(* IEC 61131-3 sources: plc-st-coding-agent/progress/evidence/f14_v14_remaining_20261113/jobs/codex_minimax-m27 (part 6) *)

(* ---- self-hard-07.candidate_01.st ---- *)
FUNCTION_BLOCK FB
VAR_INPUT
    mode                : INT;
    resetBtn            : BOOL;
    scanSeconds         : REAL;
    tempSP              : REAL;
    tempPV              : REAL;
    flowPV              : REAL;
    manualFlowSP        : REAL;
    manualValve         : REAL;
END_VAR
VAR_OUTPUT
    flowSP              : REAL;
    valveCommand        : REAL;
    fault               : BOOL;
    normalMode          : BOOL;
END_VAR
VAR
    accT                : REAL := 0.0;
    accF                : REAL := 0.0;
    mode_prev           : INT := 999;
    prev_resetBtn       : BOOL := FALSE;
    first_scan          : BOOL := TRUE;
END_VAR
VAR_TEMP
    eT                  : REAL;
    eF                  : REAL;
    trial               : REAL;
    reset_rising        : BOOL;
    mode_changed        : BOOL;
END_VAR
(* ENGINEERING_CONTRACT
 * =============================================================================
 * Modes: 0=Manual(FB), 1=Auto(inner PI), 2=Cascade(both PI loops)
 * Normal operation: mode in {0,1,2}, 0 < scanSeconds <= 10.0
 * Fault: mode outside {0,1,2} OR scanSeconds <= 0 OR scanSeconds > 10
 * -----------------------------------------------------------------------------
 * Output state retention (per LTL spec):
 * - Mode switch to 2 (cascade): flowSP, valveCommand HOLD prev; normalMode=FALSE
 * - Mode switch to 0/1: flowSP=manualFlowSP, valveCommand HOLD prev; normalMode=FALSE
 * - Manual (mode=0) normal cycle: flowSP=manualFlowSP, valveCommand=manualValve
 * - Auto (mode=1) normal cycle: flowSP=manualFlowSP; valveCommand=PI(clamped)
 * - Cascade (mode=2) normal cycle: flowSP=PI(clamped), valveCommand=PI(clamped)
 * - Fault: flowSP=manualFlowSP, valveCommand=manualValve, normalMode=FALSE
 * - Reset rising edge: same as fault initialization, fault still reports truthfully
 * -----------------------------------------------------------------------------
 * Integrators (anti-windup back-calculation):
 * - accT unit: t/h; accF unit: %; both pre-set to 0 on reset/fault/first scan
 * - acc update after output limit: acc = limited_output - Kp*e
 * - On mode change to cascade, both accT and accF retain prior cycle values
 * -----------------------------------------------------------------------------
 * Timing: Ki defined per second; scanSeconds multiplied explicitly
 * Boundaries: flowSP [0,50] t/h; valveCommand [0,100] %
 * =============================================================================
 *)
(* CONTRACT_RULES [] *)

reset_rising := resetBtn AND NOT prev_resetBtn;
mode_changed := (mode <> mode_prev);

fault := (mode < 0) OR (mode > 2) OR (scanSeconds <= 0.0) OR (scanSeconds > 10.0);

IF first_scan OR reset_rising THEN
    flowSP := manualFlowSP;
    valveCommand := manualValve;
    accT := 0.0;
    accF := 0.0;
    normalMode := FALSE;
    first_scan := FALSE;
ELSIF fault THEN
    flowSP := manualFlowSP;
    valveCommand := manualValve;
    accT := 0.0;
    accF := 0.0;
    normalMode := FALSE;
ELSE
    IF mode_changed THEN
        normalMode := FALSE;
        IF mode = 2 THEN
            // Cascade: hold both outputs
            // accT, accF retained for bumpless entry
        ELSIF (mode = 0) OR (mode = 1) THEN
            flowSP := manualFlowSP;
            // valveCommand held
        END_IF;
    ELSE
        normalMode := TRUE;
        IF mode = 2 THEN
            // Outer loop PI
            eT := tempSP - tempPV;
            accT := accT + 0.2 * eT * scanSeconds;
            trial := accT + 0.2 * eT * scanSeconds;
            flowSP := 1.0 * eT + trial;
            flowSP := LIMIT(0.0, flowSP, 50.0);
            accT := flowSP - 1.0 * eT;
            // Inner loop PI
            eF := flowSP - flowPV;
            accF := accF + 0.5 * eF * scanSeconds;
            trial := accF + 0.5 * eF * scanSeconds;
            valveCommand := 2.0 * eF + trial;
            valveCommand := LIMIT(0.0, valveCommand, 100.0);
            accF := valveCommand - 2.0 * eF;
        ELSIF mode = 1 THEN
            // Auto: flowSP from manual, inner PI
            flowSP := manualFlowSP;
            eF := flowSP - flowPV;
            accF := accF + 0.5 * eF * scanSeconds;
            trial := accF + 0.5 * eF * scanSeconds;
            valveCommand := 2.0 * eF + trial;
            valveCommand := LIMIT(0.0, valveCommand, 100.0);
            accF := valveCommand - 2.0 * eF;
        ELSIF mode = 0 THEN
            // Manual
            flowSP := manualFlowSP;
            valveCommand := manualValve;
        END_IF;
    END_IF;
END_IF;

mode_prev := mode;
prev_resetBtn := resetBtn;
END_FUNCTION_BLOCK

(* ---- self-hard-07.patch_base_02.st ---- *)
FUNCTION_BLOCK FB
VAR_INPUT
    mode                : INT;
    resetBtn            : BOOL;
    scanSeconds         : REAL;
    tempSP              : REAL;
    tempPV              : REAL;
    flowPV              : REAL;
    manualFlowSP        : REAL;
    manualValve         : REAL;
END_VAR
VAR_OUTPUT
    flowSP              : REAL;
    valveCommand        : REAL;
    fault               : BOOL;
    normalMode          : BOOL;
END_VAR
VAR
    accT                : REAL := 0.0;
    accF                : REAL := 0.0;
    mode_prev           : INT := 999;
    prev_resetBtn       : BOOL := FALSE;
    first_scan          : BOOL := TRUE;
END_VAR
VAR_TEMP
    eT                  : REAL;
    eF                  : REAL;
    trial               : REAL;
    reset_rising        : BOOL;
    mode_changed        : BOOL;
END_VAR
(* ENGINEERING_CONTRACT
 * =============================================================================
 * Modes: 0=Manual(FB), 1=Auto(inner PI), 2=Cascade(both PI loops)
 * Normal operation: mode in {0,1,2}, 0 < scanSeconds <= 10.0
 * Fault: mode outside {0,1,2} OR scanSeconds <= 0 OR scanSeconds > 10
 * -----------------------------------------------------------------------------
 * Output state retention (per LTL spec):
 * - Mode switch to 2 (cascade): flowSP, valveCommand HOLD prev; normalMode=FALSE
 * - Mode switch to 0/1: flowSP=manualFlowSP, valveCommand HOLD prev; normalMode=FALSE
 * - Manual (mode=0) normal cycle: flowSP=manualFlowSP, valveCommand=manualValve
 * - Auto (mode=1) normal cycle: flowSP=manualFlowSP; valveCommand=PI(clamped)
 * - Cascade (mode=2) normal cycle: flowSP=PI(clamped), valveCommand=PI(clamped)
 * - Fault: flowSP=manualFlowSP, valveCommand=manualValve, normalMode=FALSE
 * - Reset rising edge: same as fault initialization, fault still reports truthfully
 * -----------------------------------------------------------------------------
 * Integrators (anti-windup back-calculation):
 * - accT unit: t/h; accF unit: %; both pre-set to 0 on reset/fault/first scan
 * - acc update after output limit: acc = limited_output - Kp*e
 * - On mode change to cascade, both accT and accF retain prior cycle values
 * -----------------------------------------------------------------------------
 * Timing: Ki defined per second; scanSeconds multiplied explicitly
 * Boundaries: flowSP [0,50] t/h; valveCommand [0,100] %
 * =============================================================================
 *)
(* CONTRACT_RULES [] *)

reset_rising := resetBtn AND NOT prev_resetBtn;
mode_changed := (mode <> mode_prev);

fault := (mode < 0) OR (mode > 2) OR (scanSeconds <= 0.0) OR (scanSeconds > 10.0);

IF first_scan OR reset_rising THEN
    flowSP := manualFlowSP;
    valveCommand := manualValve;
    accT := 0.0;
    accF := 0.0;
    normalMode := FALSE;
    first_scan := FALSE;
ELSIF fault THEN
    flowSP := manualFlowSP;
    valveCommand := manualValve;
    accT := 0.0;
    accF := 0.0;
    normalMode := FALSE;
ELSE
    IF mode_changed THEN
        normalMode := FALSE;
        IF mode = 2 THEN
            // Cascade: hold both outputs
            // accT, accF retained for bumpless entry
        ELSIF (mode = 0) OR (mode = 1) THEN
            flowSP := manualFlowSP;
            // valveCommand held
        END_IF;
    ELSE
        normalMode := TRUE;
        IF mode = 2 THEN
            // Outer loop PI
            eT := tempSP - tempPV;
            accT := accT + 0.2 * eT * scanSeconds;
            trial := accT + 0.2 * eT * scanSeconds;
            flowSP := 1.0 * eT + trial;
            flowSP := LIMIT(0.0, flowSP, 50.0);
            accT := flowSP - 1.0 * eT;
            // Inner loop PI
            eF := flowSP - flowPV;
            accF := accF + 0.5 * eF * scanSeconds;
            trial := accF + 0.5 * eF * scanSeconds;
            valveCommand := 2.0 * eF + trial;
            valveCommand := LIMIT(0.0, valveCommand, 100.0);
            accF := valveCommand - 2.0 * eF;
        ELSIF mode = 1 THEN
            // Auto: flowSP from manual, inner PI
            flowSP := manualFlowSP;
            eF := flowSP - flowPV;
            accF := accF + 0.5 * eF * scanSeconds;
            trial := accF + 0.5 * eF * scanSeconds;
            valveCommand := 2.0 * eF + trial;
            valveCommand := LIMIT(0.0, valveCommand, 100.0);
            accF := valveCommand - 2.0 * eF;
        ELSIF mode = 0 THEN
            // Manual
            flowSP := manualFlowSP;
            valveCommand := manualValve;
        END_IF;
    END_IF;
END_IF;

mode_prev := mode;
prev_resetBtn := resetBtn;
END_FUNCTION_BLOCK

(* ---- self-hard-07.patch_base_03.st ---- *)
FUNCTION_BLOCK FB
VAR_INPUT
    mode                : INT;
    resetBtn            : BOOL;
    scanSeconds         : REAL;
    tempSP              : REAL;
    tempPV              : REAL;
    flowPV              : REAL;
    manualFlowSP        : REAL;
    manualValve         : REAL;
END_VAR
VAR_OUTPUT
    flowSP              : REAL;
    valveCommand        : REAL;
    fault               : BOOL;
    normalMode          : BOOL;
END_VAR
VAR
    accT                : REAL := 0.0;
    accF                : REAL := 0.0;
    mode_prev           : INT := 999;
    prev_resetBtn       : BOOL := FALSE;
    first_scan          : BOOL := TRUE;
END_VAR
VAR_TEMP
    eT                  : REAL;
    eF                  : REAL;
    trial               : REAL;
    reset_rising        : BOOL;
    mode_changed        : BOOL;
END_VAR
(* ENGINEERING_CONTRACT
 * =============================================================================
 * Modes: 0=Manual(FB), 1=Auto(inner PI), 2=Cascade(both PI loops)
 * Normal operation: mode in {0,1,2}, 0 < scanSeconds <= 10.0
 * Fault: mode outside {0,1,2} OR scanSeconds <= 0 OR scanSeconds > 10
 * -----------------------------------------------------------------------------
 * Output state retention (per LTL spec):
 * - Mode switch to 2 (cascade): flowSP, valveCommand HOLD prev; normalMode=FALSE
 * - Mode switch to 0/1: flowSP=manualFlowSP, valveCommand HOLD prev; normalMode=FALSE
 * - Manual (mode=0) normal cycle: flowSP=manualFlowSP, valveCommand=manualValve
 * - Auto (mode=1) normal cycle: flowSP=manualFlowSP; valveCommand=PI(clamped)
 * - Cascade (mode=2) normal cycle: flowSP=PI(clamped), valveCommand=PI(clamped)
 * - Fault: flowSP=manualFlowSP, valveCommand=manualValve, normalMode=FALSE
 * - Reset rising edge: same as fault initialization, fault still reports truthfully
 * -----------------------------------------------------------------------------
 * Integrators (anti-windup back-calculation):
 * - accT unit: t/h; accF unit: %; both pre-set to 0 on reset/fault/first scan
 * - acc update after output limit: acc = limited_output - Kp*e
 * - On mode change to cascade, both accT and accF retain prior cycle values
 * -----------------------------------------------------------------------------
 * Timing: Ki defined per second; scanSeconds multiplied explicitly
 * Boundaries: flowSP [0,50] t/h; valveCommand [0,100] %
 * =============================================================================
 *)
(* CONTRACT_RULES [] *)

reset_rising := resetBtn AND NOT prev_resetBtn;
mode_changed := (mode <> mode_prev);

fault := (mode < 0) OR (mode > 2) OR (scanSeconds <= 0.0) OR (scanSeconds > 10.0);

IF first_scan OR reset_rising THEN
    flowSP := manualFlowSP;
    valveCommand := manualValve;
    accT := 0.0;
    accF := 0.0;
    normalMode := FALSE;
    first_scan := FALSE;
ELSIF fault THEN
    flowSP := manualFlowSP;
    valveCommand := manualValve;
    accT := 0.0;
    accF := 0.0;
    normalMode := FALSE;
ELSE
    IF mode_changed THEN
        normalMode := FALSE;
        IF mode = 2 THEN
            // Cascade: hold both outputs
            // accT, accF retained for bumpless entry
        ELSIF (mode = 0) OR (mode = 1) THEN
            flowSP := manualFlowSP;
            // valveCommand held
        END_IF;
    ELSE
        normalMode := TRUE;
        IF mode = 2 THEN
            // Outer loop PI
            eT := tempSP - tempPV;
            accT := accT + 0.2 * eT * scanSeconds;
            trial := accT + 0.2 * eT * scanSeconds;
            flowSP := 1.0 * eT + trial;
            flowSP := LIMIT(0.0, flowSP, 50.0);
            accT := flowSP - 1.0 * eT;
            // Inner loop PI
            eF := flowSP - flowPV;
            accF := accF + 0.5 * eF * scanSeconds;
            trial := accF + 0.5 * eF * scanSeconds;
            valveCommand := 2.0 * eF + trial;
            valveCommand := LIMIT(0.0, valveCommand, 100.0);
            accF := valveCommand - 2.0 * eF;
        ELSIF mode = 1 THEN
            // Auto: flowSP from manual, inner PI
            flowSP := manualFlowSP;
            eF := flowSP - flowPV;
            accF := accF + 0.5 * eF * scanSeconds;
            trial := accF + 0.5 * eF * scanSeconds;
            valveCommand := 2.0 * eF + trial;
            valveCommand := LIMIT(0.0, valveCommand, 100.0);
            accF := valveCommand - 2.0 * eF;
        ELSIF mode = 0 THEN
            // Manual
            flowSP := manualFlowSP;
            valveCommand := manualValve;
        END_IF;
    END_IF;
END_IF;

mode_prev := mode;
prev_resetBtn := resetBtn;
END_FUNCTION_BLOCK

(* ---- self-hard-07.raw_candidate_01.st ---- *)
FUNCTION_BLOCK FB
VAR_INPUT
    mode                : INT;
    resetBtn            : BOOL;
    scanSeconds         : REAL;
    tempSP              : REAL;
    tempPV              : REAL;
    flowPV              : REAL;
    manualFlowSP        : REAL;
    manualValve         : REAL;
END_VAR
VAR_OUTPUT
    flowSP              : REAL;
    valveCommand        : REAL;
    fault               : BOOL;
    normalMode          : BOOL;
END_VAR
VAR
    accT                : REAL := 0.0;
    accF                : REAL := 0.0;
    mode_prev           : INT := 999;
    prev_resetBtn       : BOOL := FALSE;
    first_scan          : BOOL := TRUE;
END_VAR
VAR_TEMP
    eT                  : REAL;
    eF                  : REAL;
    trial               : REAL;
    reset_rising        : BOOL;
    mode_changed        : BOOL;
END_VAR
(* ENGINEERING_CONTRACT
 * =============================================================================
 * Modes: 0=Manual(FB), 1=Auto(inner PI), 2=Cascade(both PI loops)
 * Normal operation: mode in {0,1,2}, 0 < scanSeconds <= 10.0
 * Fault: mode outside {0,1,2} OR scanSeconds <= 0 OR scanSeconds > 10
 * -----------------------------------------------------------------------------
 * Output state retention (per LTL spec):
 * - Mode switch to 2 (cascade): flowSP, valveCommand HOLD prev; normalMode=FALSE
 * - Mode switch to 0/1: flowSP=manualFlowSP, valveCommand HOLD prev; normalMode=FALSE
 * - Manual (mode=0) normal cycle: flowSP=manualFlowSP, valveCommand=manualValve
 * - Auto (mode=1) normal cycle: flowSP=manualFlowSP; valveCommand=PI(clamped)
 * - Cascade (mode=2) normal cycle: flowSP=PI(clamped), valveCommand=PI(clamped)
 * - Fault: flowSP=manualFlowSP, valveCommand=manualValve, normalMode=FALSE
 * - Reset rising edge: same as fault initialization, fault still reports truthfully
 * -----------------------------------------------------------------------------
 * Integrators (anti-windup back-calculation):
 * - accT unit: t/h; accF unit: %; both pre-set to 0 on reset/fault/first scan
 * - acc update after output limit: acc = limited_output - Kp*e
 * - On mode change to cascade, both accT and accF retain prior cycle values
 * -----------------------------------------------------------------------------
 * Timing: Ki defined per second; scanSeconds multiplied explicitly
 * Boundaries: flowSP [0,50] t/h; valveCommand [0,100] %
 * =============================================================================
 *)
(* CONTRACT_RULES [] *)

reset_rising := resetBtn AND NOT prev_resetBtn;
mode_changed := (mode <> mode_prev);

fault := (mode < 0) OR (mode > 2) OR (scanSeconds <= 0.0) OR (scanSeconds > 10.0);

IF first_scan OR reset_rising THEN
    flowSP := manualFlowSP;
    valveCommand := manualValve;
    accT := 0.0;
    accF := 0.0;
    normalMode := FALSE;
    first_scan := FALSE;
ELSIF fault THEN
    flowSP := manualFlowSP;
    valveCommand := manualValve;
    accT := 0.0;
    accF := 0.0;
    normalMode := FALSE;
ELSE
    IF mode_changed THEN
        normalMode := FALSE;
        IF mode = 2 THEN
            // Cascade: hold both outputs
            // accT, accF retained for bumpless entry
        ELSIF (mode = 0) OR (mode = 1) THEN
            flowSP := manualFlowSP;
            // valveCommand held
        END_IF;
    ELSE
        normalMode := TRUE;
        IF mode = 2 THEN
            // Outer loop PI
            eT := tempSP - tempPV;
            accT := accT + 0.2 * eT * scanSeconds;
            trial := accT + 0.2 * eT * scanSeconds;
            flowSP := 1.0 * eT + trial;
            flowSP := LIMIT(0.0, flowSP, 50.0);
            accT := flowSP - 1.0 * eT;
            // Inner loop PI
            eF := flowSP - flowPV;
            accF := accF + 0.5 * eF * scanSeconds;
            trial := accF + 0.5 * eF * scanSeconds;
            valveCommand := 2.0 * eF + trial;
            valveCommand := LIMIT(0.0, valveCommand, 100.0);
            accF := valveCommand - 2.0 * eF;
        ELSIF mode = 1 THEN
            // Auto: flowSP from manual, inner PI
            flowSP := manualFlowSP;
            eF := flowSP - flowPV;
            accF := accF + 0.5 * eF * scanSeconds;
            trial := accF + 0.5 * eF * scanSeconds;
            valveCommand := 2.0 * eF + trial;
            valveCommand := LIMIT(0.0, valveCommand, 100.0);
            accF := valveCommand - 2.0 * eF;
        ELSIF mode = 0 THEN
            // Manual
            flowSP := manualFlowSP;
            valveCommand := manualValve;
        END_IF;
    END_IF;
END_IF;

mode_prev := mode;
prev_resetBtn := resetBtn;
END_FUNCTION_BLOCK

(* ---- self-medium-01.candidate_01.st ---- *)
(*
ENGINEERING_CONTRACT
================================================================================
PUB001  | Activation      : loadTrig.Q & NOT running & valid slot bounds
PUB002  | Deactivation    : loadTrig.Q & NOT running & invalid bounds/slot/content
PUB003  | Retention       : running OR NOT loadTrig.Q → valid,loadedID held
PUB004  | Same-scan order : edge detection → bounds check → slot access → latch
PUB006  | Boundary        : selSlot < 1 | selSlot > 8 → valid=FALSE, loadedID=0
PUB007  | Ratio bounds    : totalRatio < 99.0 | > 101.0 → invalid
PUB008  | Temp bounds     : temperature < 30.0 | > 180.0 → invalid
PUB009  | Content check   : recipeID = 0 → slot empty → invalid
PUB010  | Units           : REAL literals for bounds (inclusive)
PUB013  | Rising edge     : R_TRIG detects loadCmd 0→1 transition
N10-S4  | Production hold : running → loadedID = prev(loadedID)
N10-S9  | No-edge hold    : NOT loadTrig.Q → loadedID = prev(loadedID)
================================================================================
*)
(* CONTRACT_RULES [] *)

FUNCTION_BLOCK FB
VAR_INPUT
    recipe    : ARRAY[1..8] OF ST_Recipe;
    selSlot   : INT;
    loadCmd   : BOOL;
    running   : BOOL;
END_VAR

VAR_OUTPUT
    valid     : BOOL;
    loadedID  : INT;
END_VAR

VAR
    loadTrig  : R_TRIG;
END_VAR

loadTrig(CLK := loadCmd);

IF loadTrig.Q AND NOT running THEN
    IF selSlot >= 1 AND selSlot <= 8 THEN
        valid := (recipe[selSlot].recipeID <> 0)
              AND (recipe[selSlot].totalRatio >= 99.0)
              AND (recipe[selSlot].totalRatio <= 101.0)
              AND (recipe[selSlot].temperature >= 30.0)
              AND (recipe[selSlot].temperature <= 180.0);

        IF valid THEN
            loadedID := recipe[selSlot].recipeID;
        ELSE
            loadedID := 0;
        END_IF;
    ELSE
        valid    := FALSE;
        loadedID := 0;
    END_IF;
ELSE
    IF NOT loadTrig.Q AND NOT running THEN
        ; // Retain valid, loadedID
    END_IF;
END_IF;

IF running THEN
    ; // Retain valid, loadedID
END_IF;

END_FUNCTION_BLOCK

(* ---- self-medium-01.candidate_02.st ---- *)
(*
ENGINEERING_CONTRACT
================================================================================
PUB001  | Activation      : loadTrig.Q & NOT running & valid slot bounds
PUB002  | Deactivation    : loadTrig.Q & NOT running & invalid bounds/slot/content
PUB003  | Retention       : running OR NOT loadTrig.Q → valid,loadedID held
PUB004  | Same-scan order : edge detection → bounds check → slot access → latch
PUB006  | Boundary        : selSlot < 1 | selSlot > 8 → valid=FALSE, loadedID=0
PUB007  | Ratio bounds    : totalRatio < 99.0 | > 101.0 → invalid
PUB008  | Temp bounds     : temperature < 30.0 | > 180.0 → invalid
PUB009  | Content check   : recipeID = 0 → slot empty → invalid
PUB010  | Units           : REAL literals for bounds (inclusive)
PUB013  | Rising edge     : R_TRIG detects loadCmd 0→1 transition
N10-S4  | Production hold : running → loadedID = prev(loadedID)
N10-S9  | No-edge hold    : NOT loadTrig.Q → loadedID = prev(loadedID)
================================================================================
*)
(* CONTRACT_RULES [] *)

TYPE ST_Recipe :
STRUCT
    recipeID    : INT;
    totalRatio  : REAL;
    temperature : REAL;
END_STRUCT
END_TYPE;

FUNCTION_BLOCK FB
VAR_INPUT
    recipe    : ARRAY[1..8] OF ST_Recipe;
    selSlot   : INT;
    loadCmd   : BOOL;
    running   : BOOL;
END_VAR

VAR_OUTPUT
    valid     : BOOL;
    loadedID  : INT;
END_VAR

VAR
    loadTrig  : R_TRIG;
END_VAR

loadTrig(CLK := loadCmd);

IF loadTrig.Q AND NOT running THEN
    IF selSlot >= 1 AND selSlot <= 8 THEN
        valid := (recipe[selSlot].recipeID <> 0)
              AND (recipe[selSlot].totalRatio >= 99.0)
              AND (recipe[selSlot].totalRatio <= 101.0)
              AND (recipe[selSlot].temperature >= 30.0)
              AND (recipe[selSlot].temperature <= 180.0);

        IF valid THEN
            loadedID := recipe[selSlot].recipeID;
        ELSE
            loadedID := 0;
        END_IF;
    ELSE
        valid    := FALSE;
        loadedID := 0;
    END_IF;
ELSE
    IF NOT loadTrig.Q AND NOT running THEN
        ; // Retain valid, loadedID
    END_IF;
END_IF;

IF running THEN
    ; // Retain valid, loadedID
END_IF;

END_FUNCTION_BLOCK

(* ---- self-medium-01.patch_base_02.st ---- *)
(*
ENGINEERING_CONTRACT
================================================================================
PUB001  | Activation      : loadTrig.Q & NOT running & valid slot bounds
PUB002  | Deactivation    : loadTrig.Q & NOT running & invalid bounds/slot/content
PUB003  | Retention       : running OR NOT loadTrig.Q → valid,loadedID held
PUB004  | Same-scan order : edge detection → bounds check → slot access → latch
PUB006  | Boundary        : selSlot < 1 | selSlot > 8 → valid=FALSE, loadedID=0
PUB007  | Ratio bounds    : totalRatio < 99.0 | > 101.0 → invalid
PUB008  | Temp bounds     : temperature < 30.0 | > 180.0 → invalid
PUB009  | Content check   : recipeID = 0 → slot empty → invalid
PUB010  | Units           : REAL literals for bounds (inclusive)
PUB013  | Rising edge     : R_TRIG detects loadCmd 0→1 transition
N10-S4  | Production hold : running → loadedID = prev(loadedID)
N10-S9  | No-edge hold    : NOT loadTrig.Q → loadedID = prev(loadedID)
================================================================================
*)
(* CONTRACT_RULES [] *)

FUNCTION_BLOCK FB
VAR_INPUT
    recipe    : ARRAY[1..8] OF ST_Recipe;
    selSlot   : INT;
    loadCmd   : BOOL;
    running   : BOOL;
END_VAR

VAR_OUTPUT
    valid     : BOOL;
    loadedID  : INT;
END_VAR

VAR
    loadTrig  : R_TRIG;
END_VAR

loadTrig(CLK := loadCmd);

IF loadTrig.Q AND NOT running THEN
    IF selSlot >= 1 AND selSlot <= 8 THEN
        valid := (recipe[selSlot].recipeID <> 0)
              AND (recipe[selSlot].totalRatio >= 99.0)
              AND (recipe[selSlot].totalRatio <= 101.0)
              AND (recipe[selSlot].temperature >= 30.0)
              AND (recipe[selSlot].temperature <= 180.0);

        IF valid THEN
            loadedID := recipe[selSlot].recipeID;
        ELSE
            loadedID := 0;
        END_IF;
    ELSE
        valid    := FALSE;
        loadedID := 0;
    END_IF;
ELSE
    IF NOT loadTrig.Q AND NOT running THEN
        ; // Retain valid, loadedID
    END_IF;
END_IF;

IF running THEN
    ; // Retain valid, loadedID
END_IF;

END_FUNCTION_BLOCK

(* ---- self-medium-01.raw_candidate_01.st ---- *)
(*
ENGINEERING_CONTRACT
================================================================================
PUB001  | Activation      : loadTrig.Q & NOT running & valid slot bounds
PUB002  | Deactivation    : loadTrig.Q & NOT running & invalid bounds/slot/content
PUB003  | Retention       : running OR NOT loadTrig.Q → valid,loadedID held
PUB004  | Same-scan order : edge detection → bounds check → slot access → latch
PUB006  | Boundary        : selSlot < 1 | selSlot > 8 → valid=FALSE, loadedID=0
PUB007  | Ratio bounds    : totalRatio < 99.0 | > 101.0 → invalid
PUB008  | Temp bounds     : temperature < 30.0 | > 180.0 → invalid
PUB009  | Content check   : recipeID = 0 → slot empty → invalid
PUB010  | Units           : REAL literals for bounds (inclusive)
PUB013  | Rising edge     : R_TRIG detects loadCmd 0→1 transition
N10-S4  | Production hold : running → loadedID = prev(loadedID)
N10-S9  | No-edge hold    : NOT loadTrig.Q → loadedID = prev(loadedID)
================================================================================
*)
(* CONTRACT_RULES [] *)

FUNCTION_BLOCK FB
VAR_INPUT
    recipe    : ARRAY[1..8] OF ST_Recipe;
    selSlot   : INT;
    loadCmd   : BOOL;
    running   : BOOL;
END_VAR

VAR_OUTPUT
    valid     : BOOL;
    loadedID  : INT;
END_VAR

VAR
    loadTrig  : R_TRIG;
END_VAR

loadTrig(CLK := loadCmd);

IF loadTrig.Q AND NOT running THEN
    IF selSlot >= 1 AND selSlot <= 8 THEN
        valid := (recipe[selSlot].recipeID <> 0)
              AND (recipe[selSlot].totalRatio >= 99.0)
              AND (recipe[selSlot].totalRatio <= 101.0)
              AND (recipe[selSlot].temperature >= 30.0)
              AND (recipe[selSlot].temperature <= 180.0);

        IF valid THEN
            loadedID := recipe[selSlot].recipeID;
        ELSE
            loadedID := 0;
        END_IF;
    ELSE
        valid    := FALSE;
        loadedID := 0;
    END_IF;
ELSE
    IF NOT loadTrig.Q AND NOT running THEN
        ; // Retain valid, loadedID
    END_IF;
END_IF;

IF running THEN
    ; // Retain valid, loadedID
END_IF;

END_FUNCTION_BLOCK

(* ---- self-medium-01.raw_candidate_02.st ---- *)
(*
ENGINEERING_CONTRACT
================================================================================
PUB001  | Activation      : loadTrig.Q & NOT running & valid slot bounds
PUB002  | Deactivation    : loadTrig.Q & NOT running & invalid bounds/slot/content
PUB003  | Retention       : running OR NOT loadTrig.Q → valid,loadedID held
PUB004  | Same-scan order : edge detection → bounds check → slot access → latch
PUB006  | Boundary        : selSlot < 1 | selSlot > 8 → valid=FALSE, loadedID=0
PUB007  | Ratio bounds    : totalRatio < 99.0 | > 101.0 → invalid
PUB008  | Temp bounds     : temperature < 30.0 | > 180.0 → invalid
PUB009  | Content check   : recipeID = 0 → slot empty → invalid
PUB010  | Units           : REAL literals for bounds (inclusive)
PUB013  | Rising edge     : R_TRIG detects loadCmd 0→1 transition
N10-S4  | Production hold : running → loadedID = prev(loadedID)
N10-S9  | No-edge hold    : NOT loadTrig.Q → loadedID = prev(loadedID)
================================================================================
*)
(* CONTRACT_RULES [] *)

TYPE ST_Recipe :
STRUCT
    recipeID    : INT;
    totalRatio  : REAL;
    temperature : REAL;
END_STRUCT
END_TYPE

FUNCTION_BLOCK FB
VAR_INPUT
    recipe    : ARRAY[1..8] OF ST_Recipe;
    selSlot   : INT;
    loadCmd   : BOOL;
    running   : BOOL;
END_VAR

VAR_OUTPUT
    valid     : BOOL;
    loadedID  : INT;
END_VAR

VAR
    loadTrig  : R_TRIG;
END_VAR

loadTrig(CLK := loadCmd);

IF loadTrig.Q AND NOT running THEN
    IF selSlot >= 1 AND selSlot <= 8 THEN
        valid := (recipe[selSlot].recipeID <> 0)
              AND (recipe[selSlot].totalRatio >= 99.0)
              AND (recipe[selSlot].totalRatio <= 101.0)
              AND (recipe[selSlot].temperature >= 30.0)
              AND (recipe[selSlot].temperature <= 180.0);

        IF valid THEN
            loadedID := recipe[selSlot].recipeID;
        ELSE
            loadedID := 0;
        END_IF;
    ELSE
        valid    := FALSE;
        loadedID := 0;
    END_IF;
ELSE
    IF NOT loadTrig.Q AND NOT running THEN
        ; // Retain valid, loadedID
    END_IF;
END_IF;

IF running THEN
    ; // Retain valid, loadedID
END_IF;

END_FUNCTION_BLOCK

(* ---- self-medium-02.candidate_01.st ---- *)
(* ENGINEERING_CONTRACT
 * Pub: PUB001-006, PUB008-012, PUB015, PUB017, PUB019-022, PUB024-026, PUB028-038
 * Block: FB (8-point moving average with FIFO eviction)
 *
 * | Output/State     | Activation         | Retention                    | Reset/Deactivation         | Priority | Units        |
 * |------------------|--------------------|------------------------------|-----------------------------|----------|--------------|
 * | filteredValue    | Each enable scan   | Hold last when enable=FALSE  | None (retention required)   | Same-scan| REAL         |
 * | windowFull       | sampleCount=8      | Hold TRUE when full          | Clear on enable=FALSE       | Same-scan| BOOL         |
 * | sampleCount      | +1 per sample<8    | Reset to 0 when enable=FALSE | Clear on enable=FALSE       | Same-scan| INT [0..8]   |
 * | buffer/sum/idx   | Fresh start on enable| Not exposed externally      | Clear on enable=FALSE       | N/A      | VAR statics  |
 *
 * CONTRACT_RULES []
 *)
FUNCTION_BLOCK FB
VAR_INPUT
    enable    : BOOL;
    rawValue  : REAL;
END_VAR
VAR_OUTPUT
    filteredValue : REAL;
    windowFull    : BOOL;
    sampleCount   : INT;
END_VAR
VAR
    buffer     : ARRAY[0..7] OF REAL := (0,0,0,0,0,0,0,0);
    writeIndex : INT := 0;
    sum        : REAL := 0.0;
END_VAR

IF enable THEN
    (* Fresh start on transition from disabled *)
    IF sampleCount = 0 THEN
        buffer[0] := rawValue;
        buffer[1] := 0.0; buffer[2] := 0.0; buffer[3] := 0.0;
        buffer[4] := 0.0; buffer[5] := 0.0; buffer[6] := 0.0; buffer[7] := 0.0;
        writeIndex := 1;
        sum := rawValue;
        sampleCount := 1;
        filteredValue := rawValue;
        windowFull := FALSE;
    ELSE
        (* Normal operation *)
        IF sampleCount < 8 THEN
            buffer[writeIndex] := rawValue;
            sum := sum + rawValue;
            writeIndex := (writeIndex + 1) MOD 8;
            sampleCount := sampleCount + 1;
        ELSE
            (* FIFO eviction when full *)
            sum := sum - buffer[writeIndex];
            buffer[writeIndex] := rawValue;
            writeIndex := (writeIndex + 1) MOD 8;
        END_IF;
        filteredValue := sum / INT_TO_REAL(sampleCount);
        IF sampleCount >= 8 THEN
            windowFull := TRUE;
        END_IF;
    END_IF;
ELSE
    sampleCount := 0;
    windowFull := FALSE;
END_IF;

END_FUNCTION_BLOCK

(* ---- self-medium-02.candidate_02.st ---- *)
(* ENGINEERING_CONTRACT
 * Pub: PUB001-006, PUB008-012, PUB015, PUB017, PUB019-022, PUB024-026, PUB028-038
 * Block: FB (8-point moving average with FIFO eviction)
 *
 * | Output/State     | Activation         | Retention                    | Reset/Deactivation         | Priority | Units        |
 * |------------------|--------------------|------------------------------|-----------------------------|----------|--------------|
 * | filteredValue    | Each enable scan   | Hold last when enable=FALSE  | None (retention required)   | Same-scan| REAL         |
 * | windowFull       | sampleCount=8      | Hold TRUE when full          | Clear on enable=FALSE       | Same-scan| BOOL         |
 * | sampleCount      | +1 per sample<8    | Reset to 0 when enable=FALSE | Clear on enable=FALSE       | Same-scan| INT [0..8]   |
 * | buffer/sum/idx   | Fresh start on enable| Not exposed externally      | Clear on enable=FALSE       | N/A      | VAR statics  |
 *
 * CONTRACT_RULES []
 *)
FUNCTION_BLOCK FB
VAR_INPUT
    enable    : BOOL;
    rawValue  : REAL;
END_VAR
VAR_OUTPUT
    filteredValue : REAL;
    windowFull    : BOOL;
    sampleCount   : INT;
END_VAR
VAR
    buffer     : ARRAY[0..7] OF REAL := [0.0, 0.0, 0.0, 0.0, 0.0, 0.0, 0.0, 0.0];
    writeIndex : INT := 0;
    sum        : REAL := 0.0;
END_VAR

IF enable THEN
    (* Fresh start on transition from disabled *)
    IF sampleCount = 0 THEN
        buffer[0] := rawValue;
        buffer[1] := 0.0; buffer[2] := 0.0; buffer[3] := 0.0;
        buffer[4] := 0.0; buffer[5] := 0.0; buffer[6] := 0.0; buffer[7] := 0.0;
        writeIndex := 1;
        sum := rawValue;
        sampleCount := 1;
        filteredValue := rawValue;
        windowFull := FALSE;
    ELSE
        (* Normal operation *)
        IF sampleCount < 8 THEN
            buffer[writeIndex] := rawValue;
            sum := sum + rawValue;
            writeIndex := (writeIndex + 1) MOD 8;
            sampleCount := sampleCount + 1;
        ELSE
            (* FIFO eviction when full *)
            sum := sum - buffer[writeIndex];
            buffer[writeIndex] := rawValue;
            writeIndex := (writeIndex + 1) MOD 8;
        END_IF;
        filteredValue := sum / INT_TO_REAL(sampleCount);
        IF sampleCount >= 8 THEN
            windowFull := TRUE;
        END_IF;
    END_IF;
ELSE
    sampleCount := 0;
    windowFull := FALSE;
END_IF;

END_FUNCTION_BLOCK

(* ---- self-medium-02.patch_base_02.st ---- *)
(* ENGINEERING_CONTRACT
 * Pub: PUB001-006, PUB008-012, PUB015, PUB017, PUB019-022, PUB024-026, PUB028-038
 * Block: FB (8-point moving average with FIFO eviction)
 *
 * | Output/State     | Activation         | Retention                    | Reset/Deactivation         | Priority | Units        |
 * |------------------|--------------------|------------------------------|-----------------------------|----------|--------------|
 * | filteredValue    | Each enable scan   | Hold last when enable=FALSE  | None (retention required)   | Same-scan| REAL         |
 * | windowFull       | sampleCount=8      | Hold TRUE when full          | Clear on enable=FALSE       | Same-scan| BOOL         |
 * | sampleCount      | +1 per sample<8    | Reset to 0 when enable=FALSE | Clear on enable=FALSE       | Same-scan| INT [0..8]   |
 * | buffer/sum/idx   | Fresh start on enable| Not exposed externally      | Clear on enable=FALSE       | N/A      | VAR statics  |
 *
 * CONTRACT_RULES []
 *)
FUNCTION_BLOCK FB
VAR_INPUT
    enable    : BOOL;
    rawValue  : REAL;
END_VAR
VAR_OUTPUT
    filteredValue : REAL;
    windowFull    : BOOL;
    sampleCount   : INT;
END_VAR
VAR
    buffer     : ARRAY[0..7] OF REAL := (0,0,0,0,0,0,0,0);
    writeIndex : INT := 0;
    sum        : REAL := 0.0;
END_VAR

IF enable THEN
    (* Fresh start on transition from disabled *)
    IF sampleCount = 0 THEN
        buffer[0] := rawValue;
        buffer[1] := 0.0; buffer[2] := 0.0; buffer[3] := 0.0;
        buffer[4] := 0.0; buffer[5] := 0.0; buffer[6] := 0.0; buffer[7] := 0.0;
        writeIndex := 1;
        sum := rawValue;
        sampleCount := 1;
        filteredValue := rawValue;
        windowFull := FALSE;
    ELSE
        (* Normal operation *)
        IF sampleCount < 8 THEN
            buffer[writeIndex] := rawValue;
            sum := sum + rawValue;
            writeIndex := (writeIndex + 1) MOD 8;
            sampleCount := sampleCount + 1;
        ELSE
            (* FIFO eviction when full *)
            sum := sum - buffer[writeIndex];
            buffer[writeIndex] := rawValue;
            writeIndex := (writeIndex + 1) MOD 8;
        END_IF;
        filteredValue := sum / INT_TO_REAL(sampleCount);
        IF sampleCount >= 8 THEN
            windowFull := TRUE;
        END_IF;
    END_IF;
ELSE
    sampleCount := 0;
    windowFull := FALSE;
END_IF;

END_FUNCTION_BLOCK

(* ---- self-medium-02.raw_candidate_01.st ---- *)
(* ENGINEERING_CONTRACT
 * Pub: PUB001-006, PUB008-012, PUB015, PUB017, PUB019-022, PUB024-026, PUB028-038
 * Block: FB (8-point moving average with FIFO eviction)
 *
 * | Output/State     | Activation         | Retention                    | Reset/Deactivation         | Priority | Units        |
 * |------------------|--------------------|------------------------------|-----------------------------|----------|--------------|
 * | filteredValue    | Each enable scan   | Hold last when enable=FALSE  | None (retention required)   | Same-scan| REAL         |
 * | windowFull       | sampleCount=8      | Hold TRUE when full          | Clear on enable=FALSE       | Same-scan| BOOL         |
 * | sampleCount      | +1 per sample<8    | Reset to 0 when enable=FALSE | Clear on enable=FALSE       | Same-scan| INT [0..8]   |
 * | buffer/sum/idx   | Fresh start on enable| Not exposed externally      | Clear on enable=FALSE       | N/A      | VAR statics  |
 *
 * CONTRACT_RULES []
 *)
FUNCTION_BLOCK FB
VAR_INPUT
    enable    : BOOL;
    rawValue  : REAL;
END_VAR
VAR_OUTPUT
    filteredValue : REAL;
    windowFull    : BOOL;
    sampleCount   : INT;
END_VAR
VAR
    buffer     : ARRAY[0..7] OF REAL := (0,0,0,0,0,0,0,0);
    writeIndex : INT := 0;
    sum        : REAL := 0.0;
END_VAR

IF enable THEN
    (* Fresh start on transition from disabled *)
    IF sampleCount = 0 THEN
        buffer[0] := rawValue;
        buffer[1] := 0.0; buffer[2] := 0.0; buffer[3] := 0.0;
        buffer[4] := 0.0; buffer[5] := 0.0; buffer[6] := 0.0; buffer[7] := 0.0;
        writeIndex := 1;
        sum := rawValue;
        sampleCount := 1;
        filteredValue := rawValue;
        windowFull := FALSE;
    ELSE
        (* Normal operation *)
        IF sampleCount < 8 THEN
            buffer[writeIndex] := rawValue;
            sum := sum + rawValue;
            writeIndex := (writeIndex + 1) MOD 8;
            sampleCount := sampleCount + 1;
        ELSE
            (* FIFO eviction when full *)
            sum := sum - buffer[writeIndex];
            buffer[writeIndex] := rawValue;
            writeIndex := (writeIndex + 1) MOD 8;
        END_IF;
        filteredValue := sum / INT_TO_REAL(sampleCount);
        IF sampleCount >= 8 THEN
            windowFull := TRUE;
        END_IF;
    END_IF;
ELSE
    sampleCount := 0;
    windowFull := FALSE;
END_IF;

END_FUNCTION_BLOCK

(* ---- self-medium-02.raw_candidate_02.st ---- *)
(* ENGINEERING_CONTRACT
 * Pub: PUB001-006, PUB008-012, PUB015, PUB017, PUB019-022, PUB024-026, PUB028-038
 * Block: FB (8-point moving average with FIFO eviction)
 *
 * | Output/State     | Activation         | Retention                    | Reset/Deactivation         | Priority | Units        |
 * |------------------|--------------------|------------------------------|-----------------------------|----------|--------------|
 * | filteredValue    | Each enable scan   | Hold last when enable=FALSE  | None (retention required)   | Same-scan| REAL         |
 * | windowFull       | sampleCount=8      | Hold TRUE when full          | Clear on enable=FALSE       | Same-scan| BOOL         |
 * | sampleCount      | +1 per sample<8    | Reset to 0 when enable=FALSE | Clear on enable=FALSE       | Same-scan| INT [0..8]   |
 * | buffer/sum/idx   | Fresh start on enable| Not exposed externally      | Clear on enable=FALSE       | N/A      | VAR statics  |
 *
 * CONTRACT_RULES []
 *)
FUNCTION_BLOCK FB
VAR_INPUT
    enable    : BOOL;
    rawValue  : REAL;
END_VAR
VAR_OUTPUT
    filteredValue : REAL;
    windowFull    : BOOL;
    sampleCount   : INT;
END_VAR
VAR
    buffer     : ARRAY[0..7] OF REAL := [0.0, 0.0, 0.0, 0.0, 0.0, 0.0, 0.0, 0.0];
    writeIndex : INT := 0;
    sum        : REAL := 0.0;
END_VAR

IF enable THEN
    (* Fresh start on transition from disabled *)
    IF sampleCount = 0 THEN
        buffer[0] := rawValue;
        buffer[1] := 0.0; buffer[2] := 0.0; buffer[3] := 0.0;
        buffer[4] := 0.0; buffer[5] := 0.0; buffer[6] := 0.0; buffer[7] := 0.0;
        writeIndex := 1;
        sum := rawValue;
        sampleCount := 1;
        filteredValue := rawValue;
        windowFull := FALSE;
    ELSE
        (* Normal operation *)
        IF sampleCount < 8 THEN
            buffer[writeIndex] := rawValue;
            sum := sum + rawValue;
            writeIndex := (writeIndex + 1) MOD 8;
            sampleCount := sampleCount + 1;
        ELSE
            (* FIFO eviction when full *)
            sum := sum - buffer[writeIndex];
            buffer[writeIndex] := rawValue;
            writeIndex := (writeIndex + 1) MOD 8;
        END_IF;
        filteredValue := sum / INT_TO_REAL(sampleCount);
        IF sampleCount >= 8 THEN
            windowFull := TRUE;
        END_IF;
    END_IF;
ELSE
    sampleCount := 0;
    windowFull := FALSE;
END_IF;

END_FUNCTION_BLOCK

(* ---- self-medium-03.candidate_01.st ---- *)
// ENGINEERING_CONTRACT
// Pub IDs | Activation           | Retention                 | Explicit Reset           | Same-scan Priority | Units
// --------|----------------------|---------------------------|--------------------------|--------------------|------
// motorUp | Rising openBtn in    | Run until openLimit or    | obstacle->stop, reset->  | obstacle > limits  | BOOL
//         | IDLE, no obstacle,   | obstacle, stays latched   | stop, other outputs off  | > new start        |
//         | closeBtn=FALSE,      | during fault              |                          |                    |
//         | !openLimit           |                           |                          |                    |
// --------|----------------------|---------------------------|--------------------------|--------------------|------
// motorDown| Rising closeBtn in  | Run until closeLimit or   | obstacle->stop, reset->  | obstacle > limits  | BOOL
//         | IDLE, no obstacle,   | obstacle, stays latched   | stop, other outputs off  | > new start        |
//         | openBtn=FALSE,       | during fault              |                          |                    |
//         | !closeLimit          |                           |                          |                    |
// --------|----------------------|---------------------------|--------------------------|--------------------|------
// errorFlag| obstacle in any     | Latch until valid reset   | reset: no obstacle AND   | always highest     | BOOL
//         | state                | (requires no obstacle     | rising bothBtns          | priority           |
//         |                      | AND rising bothBtns)      |                          |                    |
// --------|----------------------|---------------------------|--------------------------|--------------------|------
// CONTRACT_RULES [{"kind":"hold_until_reset","output":"errorFlag","set_input":"obstacle","reset_input":"risingBothBtn"}]

FUNCTION_BLOCK FB
VAR_INPUT
    openBtn    : BOOL;
    closeBtn   : BOOL;
    openLimit  : BOOL;
    closeLimit : BOOL;
    obstacle   : BOOL;
END_VAR
VAR_OUTPUT
    motorUp    : BOOL;
    motorDown  : BOOL;
    errorFlag  : BOOL;
END_VAR
VAR
    state        : INT; // 0=IDLE, 1=OPENING, 2=CLOSING, 3=FAULT
    prevOpenBtn  : BOOL;
    prevCloseBtn : BOOL;
    prevObstacle : BOOL;
    prevErrorFlag: BOOL;
    bothHeldPrev : BOOL;
END_VAR
VAR
    risingOpenBtn  : BOOL;
    risingCloseBtn : BOOL;
    risingBothBtn  : BOOL;
END_VAR

    // Rising edge detection
    risingOpenBtn  := openBtn AND NOT prevOpenBtn;
    risingCloseBtn := closeBtn AND NOT prevCloseBtn;
    risingBothBtn  := (openBtn AND closeBtn) AND NOT bothHeldPrev;

    // ---- Priority 1: Obstacle handling ----
    IF obstacle THEN
        motorUp   := FALSE;
        motorDown := FALSE;
        errorFlag := TRUE;
        state     := 3; // FAULT
        GOTO scan_end;
    END_IF;

    // ---- Priority 2: Fault state latching ----
    IF state = 3 THEN
        // Latched: motors off, wait for valid reset
        motorUp   := FALSE;
        motorDown := FALSE;
        // Valid reset: no obstacle AND rising both buttons
        IF risingBothBtn THEN
            errorFlag := FALSE;
            state     := 0; // IDLE
        ELSE
            errorFlag := TRUE;
        END_IF;
        GOTO scan_end;
    END_IF;

    // ---- Normal operation: IDLE, OPENING, CLOSING ----
    CASE state OF
        0: // IDLE
            motorUp   := FALSE;
            motorDown := FALSE;
            // Start opening: rising openBtn, closeBtn=FALSE, no obstacle, not at limit
            IF risingOpenBtn AND NOT closeBtn AND NOT openLimit THEN
                motorUp  := TRUE;
                motorDown:= FALSE;
                state    := 1; // OPENING
            // Start closing: rising closeBtn, openBtn=FALSE, no obstacle, not at limit
            ELSIF risingCloseBtn AND NOT openBtn AND NOT closeLimit THEN
                motorUp   := FALSE;
                motorDown := TRUE;
                state     := 2; // CLOSING
            END_IF;

        1: // OPENING
            motorUp   := TRUE;
            motorDown := FALSE;
            // Stop at open limit
            IF openLimit THEN
                motorUp  := FALSE;
                motorDown:= FALSE;
                state    := 0; // IDLE
            END_IF;

        2: // CLOSING
            motorUp   := FALSE;
            motorDown := TRUE;
            // Stop at close limit
            IF closeLimit THEN
                motorUp  := FALSE;
                motorDown:= FALSE;
                state    := 0; // IDLE
            END_IF;
    END_CASE;

scan_end:
    // Update previous inputs for next scan
    prevOpenBtn   := openBtn;
    prevCloseBtn  := closeBtn;
    prevObstacle  := obstacle;
    prevErrorFlag := errorFlag;
    bothHeldPrev  := openBtn AND closeBtn;

END_FUNCTION_BLOCK

(* ---- self-medium-03.candidate_02.st ---- *)
// ENGINEERING_CONTRACT
// Pub IDs | Activation           | Retention                 | Explicit Reset           | Same-scan Priority | Units
// --------|----------------------|---------------------------|--------------------------|--------------------|------
// motorUp | Rising openBtn in    | Run until openLimit or    | obstacle->stop, reset->  | obstacle > limits  | BOOL
//         | IDLE, no obstacle,   | obstacle, stays latched   | stop, other outputs off  | > new start        |
//         | closeBtn=FALSE,      | during fault              |                          |                    |
//         | !openLimit           |                           |                          |                    |
// --------|----------------------|---------------------------|--------------------------|--------------------|------
// motorDown| Rising closeBtn in  | Run until closeLimit or   | obstacle->stop, reset->  | obstacle > limits  | BOOL
//         | IDLE, no obstacle,   | obstacle, stays latched   | stop, other outputs off  | > new start        |
//         | openBtn=FALSE,       | during fault              |                          |                    |
//         | !closeLimit          |                           |                          |                    |
// --------|----------------------|---------------------------|--------------------------|--------------------|------
// errorFlag| obstacle in any     | Latch until valid reset   | reset: no obstacle AND   | always highest     | BOOL
//         | state                | (requires no obstacle     | rising bothBtns          | priority           |
//         |                      | AND rising bothBtns)      |                          |                    |
// --------|----------------------|---------------------------|--------------------------|--------------------|------
// CONTRACT_RULES [{"kind":"hold_until_reset","output":"errorFlag","set_input":"obstacle","reset_input":"risingBothBtn"}]

FUNCTION_BLOCK FB
VAR_INPUT
    openBtn    : BOOL;
    closeBtn   : BOOL;
    openLimit  : BOOL;
    closeLimit : BOOL;
    obstacle   : BOOL;
END_VAR
VAR_OUTPUT
    motorUp    : BOOL;
    motorDown  : BOOL;
    errorFlag  : BOOL;
END_VAR
VAR
    state        : INT; // 0=IDLE, 1=OPENING, 2=CLOSING, 3=FAULT
    prevOpenBtn  : BOOL;
    prevCloseBtn : BOOL;
    prevObstacle : BOOL;
    prevErrorFlag: BOOL;
    bothHeldPrev : BOOL;
END_VAR
VAR
    risingOpenBtn  : BOOL;
    risingCloseBtn : BOOL;
    risingBothBtn  : BOOL;
END_VAR

    // Rising edge detection
    risingOpenBtn  := openBtn AND NOT prevOpenBtn;
    risingCloseBtn := closeBtn AND NOT prevCloseBtn;
    risingBothBtn  := (openBtn AND closeBtn) AND NOT bothHeldPrev;

    // ---- Priority 1: Obstacle handling ----
    IF obstacle THEN
        motorUp   := FALSE;
        motorDown := FALSE;
        errorFlag := TRUE;
        state     := 3; // FAULT
    ELSE
        // ---- Priority 2: Fault state latching ----
        IF state = 3 THEN
            motorUp   := FALSE;
            motorDown := FALSE;
            IF risingBothBtn THEN
                errorFlag := FALSE;
                state     := 0;
            ELSE
                errorFlag := TRUE;
            END_IF;
        ELSE
            // ---- Normal operation: IDLE, OPENING, CLOSING ----
            CASE state OF
                0: // IDLE
                    motorUp   := FALSE;
                    motorDown := FALSE;
                    IF risingOpenBtn AND NOT closeBtn AND NOT openLimit THEN
                        motorUp   := TRUE;
                        motorDown := FALSE;
                        state     := 1;
                    ELSIF risingCloseBtn AND NOT openBtn AND NOT closeLimit THEN
                        motorUp   := FALSE;
                        motorDown := TRUE;
                        state     := 2;
                    END_IF;

                1: // OPENING
                    motorUp   := TRUE;
                    motorDown := FALSE;
                    IF openLimit THEN
                        motorUp   := FALSE;
                        motorDown := FALSE;
                        state     := 0;
                    END_IF;

                2: // CLOSING
                    motorUp   := FALSE;
                    motorDown := TRUE;
                    IF closeLimit THEN
                        motorUp   := FALSE;
                        motorDown := FALSE;
                        state     := 0;
                    END_IF;
            END_CASE;
        END_IF;
    END_IF;

    // Update previous inputs for next scan
    prevOpenBtn   := openBtn;
    prevCloseBtn  := closeBtn;
    prevObstacle  := obstacle;
    prevErrorFlag := errorFlag;
    bothHeldPrev  := openBtn AND closeBtn;

END_FUNCTION_BLOCK

(* ---- self-medium-03.patch_base_02.st ---- *)
// ENGINEERING_CONTRACT
// Pub IDs | Activation           | Retention                 | Explicit Reset           | Same-scan Priority | Units
// --------|----------------------|---------------------------|--------------------------|--------------------|------
// motorUp | Rising openBtn in    | Run until openLimit or    | obstacle->stop, reset->  | obstacle > limits  | BOOL
//         | IDLE, no obstacle,   | obstacle, stays latched   | stop, other outputs off  | > new start        |
//         | closeBtn=FALSE,      | during fault              |                          |                    |
//         | !openLimit           |                           |                          |                    |
// --------|----------------------|---------------------------|--------------------------|--------------------|------
// motorDown| Rising closeBtn in  | Run until closeLimit or   | obstacle->stop, reset->  | obstacle > limits  | BOOL
//         | IDLE, no obstacle,   | obstacle, stays latched   | stop, other outputs off  | > new start        |
//         | openBtn=FALSE,       | during fault              |                          |                    |
//         | !closeLimit          |                           |                          |                    |
// --------|----------------------|---------------------------|--------------------------|--------------------|------
// errorFlag| obstacle in any     | Latch until valid reset   | reset: no obstacle AND   | always highest     | BOOL
//         | state                | (requires no obstacle     | rising bothBtns          | priority           |
//         |                      | AND rising bothBtns)      |                          |                    |
// --------|----------------------|---------------------------|--------------------------|--------------------|------
// CONTRACT_RULES [{"kind":"hold_until_reset","output":"errorFlag","set_input":"obstacle","reset_input":"risingBothBtn"}]

FUNCTION_BLOCK FB
VAR_INPUT
    openBtn    : BOOL;
    closeBtn   : BOOL;
    openLimit  : BOOL;
    closeLimit : BOOL;
    obstacle   : BOOL;
END_VAR
VAR_OUTPUT
    motorUp    : BOOL;
    motorDown  : BOOL;
    errorFlag  : BOOL;
END_VAR
VAR
    state        : INT; // 0=IDLE, 1=OPENING, 2=CLOSING, 3=FAULT
    prevOpenBtn  : BOOL;
    prevCloseBtn : BOOL;
    prevObstacle : BOOL;
    prevErrorFlag: BOOL;
    bothHeldPrev : BOOL;
END_VAR
VAR
    risingOpenBtn  : BOOL;
    risingCloseBtn : BOOL;
    risingBothBtn  : BOOL;
END_VAR

    // Rising edge detection
    risingOpenBtn  := openBtn AND NOT prevOpenBtn;
    risingCloseBtn := closeBtn AND NOT prevCloseBtn;
    risingBothBtn  := (openBtn AND closeBtn) AND NOT bothHeldPrev;

    // ---- Priority 1: Obstacle handling ----
    IF obstacle THEN
        motorUp   := FALSE;
        motorDown := FALSE;
        errorFlag := TRUE;
        state     := 3; // FAULT
        GOTO scan_end;
    END_IF;

    // ---- Priority 2: Fault state latching ----
    IF state = 3 THEN
        // Latched: motors off, wait for valid reset
        motorUp   := FALSE;
        motorDown := FALSE;
        // Valid reset: no obstacle AND rising both buttons
        IF risingBothBtn THEN
            errorFlag := FALSE;
            state     := 0; // IDLE
        ELSE
            errorFlag := TRUE;
        END_IF;
        GOTO scan_end;
    END_IF;

    // ---- Normal operation: IDLE, OPENING, CLOSING ----
    CASE state OF
        0: // IDLE
            motorUp   := FALSE;
            motorDown := FALSE;
            // Start opening: rising openBtn, closeBtn=FALSE, no obstacle, not at limit
            IF risingOpenBtn AND NOT closeBtn AND NOT openLimit THEN
                motorUp  := TRUE;
                motorDown:= FALSE;
                state    := 1; // OPENING
            // Start closing: rising closeBtn, openBtn=FALSE, no obstacle, not at limit
            ELSIF risingCloseBtn AND NOT openBtn AND NOT closeLimit THEN
                motorUp   := FALSE;
                motorDown := TRUE;
                state     := 2; // CLOSING
            END_IF;

        1: // OPENING
            motorUp   := TRUE;
            motorDown := FALSE;
            // Stop at open limit
            IF openLimit THEN
                motorUp  := FALSE;
                motorDown:= FALSE;
                state    := 0; // IDLE
            END_IF;

        2: // CLOSING
            motorUp   := FALSE;
            motorDown := TRUE;
            // Stop at close limit
            IF closeLimit THEN
                motorUp  := FALSE;
                motorDown:= FALSE;
                state    := 0; // IDLE
            END_IF;
    END_CASE;

scan_end:
    // Update previous inputs for next scan
    prevOpenBtn   := openBtn;
    prevCloseBtn  := closeBtn;
    prevObstacle  := obstacle;
    prevErrorFlag := errorFlag;
    bothHeldPrev  := openBtn AND closeBtn;

END_FUNCTION_BLOCK

(* ---- self-medium-03.raw_candidate_01.st ---- *)
// ENGINEERING_CONTRACT
// Pub IDs | Activation           | Retention                 | Explicit Reset           | Same-scan Priority | Units
// --------|----------------------|---------------------------|--------------------------|--------------------|------
// motorUp | Rising openBtn in    | Run until openLimit or    | obstacle->stop, reset->  | obstacle > limits  | BOOL
//         | IDLE, no obstacle,   | obstacle, stays latched   | stop, other outputs off  | > new start        |
//         | closeBtn=FALSE,      | during fault              |                          |                    |
//         | !openLimit           |                           |                          |                    |
// --------|----------------------|---------------------------|--------------------------|--------------------|------
// motorDown| Rising closeBtn in  | Run until closeLimit or   | obstacle->stop, reset->  | obstacle > limits  | BOOL
//         | IDLE, no obstacle,   | obstacle, stays latched   | stop, other outputs off  | > new start        |
//         | openBtn=FALSE,       | during fault              |                          |                    |
//         | !closeLimit          |                           |                          |                    |
// --------|----------------------|---------------------------|--------------------------|--------------------|------
// errorFlag| obstacle in any     | Latch until valid reset   | reset: no obstacle AND   | always highest     | BOOL
//         | state                | (requires no obstacle     | rising bothBtns          | priority           |
//         |                      | AND rising bothBtns)      |                          |                    |
// --------|----------------------|---------------------------|--------------------------|--------------------|------
// CONTRACT_RULES [{"kind":"hold_until_reset","output":"errorFlag","set_input":"obstacle","reset_input":"risingBothBtn"}]

FUNCTION_BLOCK FB
VAR_INPUT
    openBtn    : BOOL;
    closeBtn   : BOOL;
    openLimit  : BOOL;
    closeLimit : BOOL;
    obstacle   : BOOL;
END_VAR
VAR_OUTPUT
    motorUp    : BOOL;
    motorDown  : BOOL;
    errorFlag  : BOOL;
END_VAR
VAR
    state        : INT; // 0=IDLE, 1=OPENING, 2=CLOSING, 3=FAULT
    prevOpenBtn  : BOOL;
    prevCloseBtn : BOOL;
    prevObstacle : BOOL;
    prevErrorFlag: BOOL;
    bothHeldPrev : BOOL;
END_VAR
VAR
    risingOpenBtn  : BOOL;
    risingCloseBtn : BOOL;
    risingBothBtn  : BOOL;
END_VAR

    // Rising edge detection
    risingOpenBtn  := openBtn AND NOT prevOpenBtn;
    risingCloseBtn := closeBtn AND NOT prevCloseBtn;
    risingBothBtn  := (openBtn AND closeBtn) AND NOT bothHeldPrev;

    // ---- Priority 1: Obstacle handling ----
    IF obstacle THEN
        motorUp   := FALSE;
        motorDown := FALSE;
        errorFlag := TRUE;
        state     := 3; // FAULT
        GOTO scan_end;
    END_IF

    // ---- Priority 2: Fault state latching ----
    IF state = 3 THEN
        // Latched: motors off, wait for valid reset
        motorUp   := FALSE;
        motorDown := FALSE;
        // Valid reset: no obstacle AND rising both buttons
        IF risingBothBtn THEN
            errorFlag := FALSE;
            state     := 0; // IDLE
        ELSE
            errorFlag := TRUE;
        END_IF
        GOTO scan_end;
    END_IF

    // ---- Normal operation: IDLE, OPENING, CLOSING ----
    CASE state OF
        0: // IDLE
            motorUp   := FALSE;
            motorDown := FALSE;
            // Start opening: rising openBtn, closeBtn=FALSE, no obstacle, not at limit
            IF risingOpenBtn AND NOT closeBtn AND NOT openLimit THEN
                motorUp  := TRUE;
                motorDown:= FALSE;
                state    := 1; // OPENING
            // Start closing: rising closeBtn, openBtn=FALSE, no obstacle, not at limit
            ELSIF risingCloseBtn AND NOT openBtn AND NOT closeLimit THEN
                motorUp   := FALSE;
                motorDown := TRUE;
                state     := 2; // CLOSING
            END_IF;

        1: // OPENING
            motorUp   := TRUE;
            motorDown := FALSE;
            // Stop at open limit
            IF openLimit THEN
                motorUp  := FALSE;
                motorDown:= FALSE;
                state    := 0; // IDLE
            END_IF;

        2: // CLOSING
            motorUp   := FALSE;
            motorDown := TRUE;
            // Stop at close limit
            IF closeLimit THEN
                motorUp  := FALSE;
                motorDown:= FALSE;
                state    := 0; // IDLE
            END_IF;
    END_CASE;

scan_end:
    // Update previous inputs for next scan
    prevOpenBtn   := openBtn;
    prevCloseBtn  := closeBtn;
    prevObstacle  := obstacle;
    prevErrorFlag := errorFlag;
    bothHeldPrev  := openBtn AND closeBtn;

END_FUNCTION_BLOCK

(* ---- self-medium-03.raw_candidate_02.st ---- *)
// ENGINEERING_CONTRACT
// Pub IDs | Activation           | Retention                 | Explicit Reset           | Same-scan Priority | Units
// --------|----------------------|---------------------------|--------------------------|--------------------|------
// motorUp | Rising openBtn in    | Run until openLimit or    | obstacle->stop, reset->  | obstacle > limits  | BOOL
//         | IDLE, no obstacle,   | obstacle, stays latched   | stop, other outputs off  | > new start        |
//         | closeBtn=FALSE,      | during fault              |                          |                    |
//         | !openLimit           |                           |                          |                    |
// --------|----------------------|---------------------------|--------------------------|--------------------|------
// motorDown| Rising closeBtn in  | Run until closeLimit or   | obstacle->stop, reset->  | obstacle > limits  | BOOL
//         | IDLE, no obstacle,   | obstacle, stays latched   | stop, other outputs off  | > new start        |
//         | openBtn=FALSE,       | during fault              |                          |                    |
//         | !closeLimit          |                           |                          |                    |
// --------|----------------------|---------------------------|--------------------------|--------------------|------
// errorFlag| obstacle in any     | Latch until valid reset   | reset: no obstacle AND   | always highest     | BOOL
//         | state                | (requires no obstacle     | rising bothBtns          | priority           |
//         |                      | AND rising bothBtns)      |                          |                    |
// --------|----------------------|---------------------------|--------------------------|--------------------|------
// CONTRACT_RULES [{"kind":"hold_until_reset","output":"errorFlag","set_input":"obstacle","reset_input":"risingBothBtn"}]

FUNCTION_BLOCK FB
VAR_INPUT
    openBtn    : BOOL;
    closeBtn   : BOOL;
    openLimit  : BOOL;
    closeLimit : BOOL;
    obstacle   : BOOL;
END_VAR
VAR_OUTPUT
    motorUp    : BOOL;
    motorDown  : BOOL;
    errorFlag  : BOOL;
END_VAR
VAR
    state        : INT; // 0=IDLE, 1=OPENING, 2=CLOSING, 3=FAULT
    prevOpenBtn  : BOOL;
    prevCloseBtn : BOOL;
    prevObstacle : BOOL;
    prevErrorFlag: BOOL;
    bothHeldPrev : BOOL;
END_VAR
VAR
    risingOpenBtn  : BOOL;
    risingCloseBtn : BOOL;
    risingBothBtn  : BOOL;
END_VAR

    // Rising edge detection
    risingOpenBtn  := openBtn AND NOT prevOpenBtn;
    risingCloseBtn := closeBtn AND NOT prevCloseBtn;
    risingBothBtn  := (openBtn AND closeBtn) AND NOT bothHeldPrev;

    // ---- Priority 1: Obstacle handling ----
    IF obstacle THEN
        motorUp   := FALSE;
        motorDown := FALSE;
        errorFlag := TRUE;
        state     := 3; // FAULT
    ELSE
        // ---- Priority 2: Fault state latching ----
        IF state = 3 THEN
            motorUp   := FALSE;
            motorDown := FALSE;
            IF risingBothBtn THEN
                errorFlag := FALSE;
                state     := 0;
            ELSE
                errorFlag := TRUE;
            END_IF;
        ELSE
            // ---- Normal operation: IDLE, OPENING, CLOSING ----
            CASE state OF
                0: // IDLE
                    motorUp   := FALSE;
                    motorDown := FALSE;
                    IF risingOpenBtn AND NOT closeBtn AND NOT openLimit THEN
                        motorUp   := TRUE;
                        motorDown := FALSE;
                        state     := 1;
                    ELSIF risingCloseBtn AND NOT openBtn AND NOT closeLimit THEN
                        motorUp   := FALSE;
                        motorDown := TRUE;
                        state     := 2;
                    END_IF;

                1: // OPENING
                    motorUp   := TRUE;
                    motorDown := FALSE;
                    IF openLimit THEN
                        motorUp   := FALSE;
                        motorDown := FALSE;
                        state     := 0;
                    END_IF;

                2: // CLOSING
                    motorUp   := FALSE;
                    motorDown := TRUE;
                    IF closeLimit THEN
                        motorUp   := FALSE;
                        motorDown := FALSE;
                        state     := 0;
                    END_IF;
            END_CASE;
        END_IF;
    END_IF;

    // Update previous inputs for next scan
    prevOpenBtn   := openBtn;
    prevCloseBtn  := closeBtn;
    prevObstacle  := obstacle;
    prevErrorFlag := errorFlag;
    bothHeldPrev  := openBtn AND closeBtn;

END_FUNCTION_BLOCK

(* ---- self-medium-04.candidate_01.st ---- *)
(* ENGINEERING_CONTRACT *)
(*
PUB001-PUB005: State machine (idle/filling/pending)
- valveOpen: active in filling, reset clears it, held until target reached
- fillsToday: monotonic up, reset to 0, saturates at 32767
- pendingConfirm: set when valve closes without immediate doneSensor, cleared on confirmation or reset

PUB006: startBtn rising edge triggers new bottle (only in idle or pending)
PUB007: resetBtn rising edge takes absolute priority, clears all state
PUB008: doneSensor level-triggered confirmation (checked after valve state set)
PUB009-PUB011: flowVol accumulated per scan in tmp_accVol; start scan includes its own flowVol
PUB012-PUB016: saturation behavior, no repeat count, no count while filling
*)
(* CONTRACT_RULES [] *)

FUNCTION_BLOCK FB
VAR_INPUT
    startBtn   : BOOL;
    resetBtn   : BOOL;
    doneSensor : BOOL;
    targetVol  : REAL;
    flowVol    : REAL;
END_VAR
VAR_OUTPUT
    valveOpen  : BOOL;
    fillsToday : INT;
END_VAR
VAR
    state           : INT;       // 0=idle, 1=filling, 2=pendingConfirm
    tmp_accVol      : REAL;      // accumulated volume for current bottle
    tmp_pending     : BOOL;      // bottle waiting for doneSensor confirmation
    prev_startBtn   : BOOL;      // previous scan startBtn (power-on FALSE)
    prev_resetBtn   : BOOL;      // previous scan resetBtn (power-on FALSE)
    tmp_risingStart : BOOL;
    tmp_risingReset : BOOL;
END_VAR

// Rising edge detection
tmp_risingStart := startBtn AND NOT prev_startBtn;
tmp_risingReset := resetBtn AND NOT prev_resetBtn;

// Update previous values
prev_startBtn := startBtn;
prev_resetBtn := resetBtn;

// State machine
IF tmp_risingReset THEN
    fillsToday := 0;
    valveOpen := FALSE;
    tmp_pending := FALSE;
    tmp_accVol := 0.0;
    state := 0;
ELSE
    CASE state OF
        0: // idle
            IF tmp_risingStart THEN
                IF tmp_pending THEN
                    tmp_pending := FALSE;
                END_IF;
                tmp_accVol := flowVol;
                IF flowVol >= targetVol THEN
                    valveOpen := FALSE;
                    tmp_pending := TRUE;
                    state := 2;
                ELSE
                    valveOpen := TRUE;
                    state := 1;
                END_IF;
            END_IF;

        1: // filling
            tmp_accVol := tmp_accVol + flowVol;
            IF tmp_accVol >= targetVol THEN
                valveOpen := FALSE;
                tmp_pending := TRUE;
                state := 2;
            END_IF;

        2: // pendingConfirm
            IF tmp_risingStart THEN
                IF tmp_pending THEN
                    tmp_pending := FALSE;
                END_IF;
                tmp_accVol := flowVol;
                IF flowVol >= targetVol THEN
                    valveOpen := FALSE;
                    tmp_pending := TRUE;
                ELSE
                    valveOpen := TRUE;
                    state := 1;
                END_IF;
            ELSIF doneSensor THEN
                IF fillsToday < 32767 THEN
                    fillsToday := fillsToday + 1;
                END_IF;
                tmp_pending := FALSE;
                state := 0;
            END_IF;
    END_CASE;
END_IF;

END_FUNCTION_BLOCK

(* ---- self-medium-04.patch_base_02.st ---- *)
(* ENGINEERING_CONTRACT *)
(*
PUB001-PUB005: State machine (idle/filling/pending)
- valveOpen: active in filling, reset clears it, held until target reached
- fillsToday: monotonic up, reset to 0, saturates at 32767
- pendingConfirm: set when valve closes without immediate doneSensor, cleared on confirmation or reset

PUB006: startBtn rising edge triggers new bottle (only in idle or pending)
PUB007: resetBtn rising edge takes absolute priority, clears all state
PUB008: doneSensor level-triggered confirmation (checked after valve state set)
PUB009-PUB011: flowVol accumulated per scan in tmp_accVol; start scan includes its own flowVol
PUB012-PUB016: saturation behavior, no repeat count, no count while filling
*)
(* CONTRACT_RULES [] *)

FUNCTION_BLOCK FB
VAR_INPUT
    startBtn   : BOOL;
    resetBtn   : BOOL;
    doneSensor : BOOL;
    targetVol  : REAL;
    flowVol    : REAL;
END_VAR
VAR_OUTPUT
    valveOpen  : BOOL;
    fillsToday : INT;
END_VAR
VAR
    state           : INT;       // 0=idle, 1=filling, 2=pendingConfirm
    tmp_accVol      : REAL;      // accumulated volume for current bottle
    tmp_pending     : BOOL;      // bottle waiting for doneSensor confirmation
    prev_startBtn   : BOOL;      // previous scan startBtn (power-on FALSE)
    prev_resetBtn   : BOOL;      // previous scan resetBtn (power-on FALSE)
    tmp_risingStart : BOOL;
    tmp_risingReset : BOOL;
END_VAR

// Rising edge detection
tmp_risingStart := startBtn AND NOT prev_startBtn;
tmp_risingReset := resetBtn AND NOT prev_resetBtn;

// Update previous values
prev_startBtn := startBtn;
prev_resetBtn := resetBtn;

// State machine
IF tmp_risingReset THEN
    fillsToday := 0;
    valveOpen := FALSE;
    tmp_pending := FALSE;
    tmp_accVol := 0.0;
    state := 0;
ELSE
    CASE state OF
        0: // idle
            IF tmp_risingStart THEN
                IF tmp_pending THEN
                    tmp_pending := FALSE;
                END_IF;
                tmp_accVol := flowVol;
                IF flowVol >= targetVol THEN
                    valveOpen := FALSE;
                    tmp_pending := TRUE;
                    state := 2;
                ELSE
                    valveOpen := TRUE;
                    state := 1;
                END_IF;
            END_IF;

        1: // filling
            tmp_accVol := tmp_accVol + flowVol;
            IF tmp_accVol >= targetVol THEN
                valveOpen := FALSE;
                tmp_pending := TRUE;
                state := 2;
            END_IF;

        2: // pendingConfirm
            IF tmp_risingStart THEN
                IF tmp_pending THEN
                    tmp_pending := FALSE;
                END_IF;
                tmp_accVol := flowVol;
                IF flowVol >= targetVol THEN
                    valveOpen := FALSE;
                    tmp_pending := TRUE;
                ELSE
                    valveOpen := TRUE;
                    state := 1;
                END_IF;
            ELSIF doneSensor THEN
                IF fillsToday < 32767 THEN
                    fillsToday := fillsToday + 1;
                END_IF;
                tmp_pending := FALSE;
                state := 0;
            END_IF;
    END_CASE;
END_IF;

END_FUNCTION_BLOCK

(* ---- self-medium-04.patch_base_03.st ---- *)
(* ENGINEERING_CONTRACT *)
(*
PUB001-PUB005: State machine (idle/filling/pending)
- valveOpen: active in filling, reset clears it, held until target reached
- fillsToday: monotonic up, reset to 0, saturates at 32767
- pendingConfirm: set when valve closes without immediate doneSensor, cleared on confirmation or reset

PUB006: startBtn rising edge triggers new bottle (only in idle or pending)
PUB007: resetBtn rising edge takes absolute priority, clears all state
PUB008: doneSensor level-triggered confirmation (checked after valve state set)
PUB009-PUB011: flowVol accumulated per scan in tmp_accVol; start scan includes its own flowVol
PUB012-PUB016: saturation behavior, no repeat count, no count while filling
*)
(* CONTRACT_RULES [] *)

FUNCTION_BLOCK FB
VAR_INPUT
    startBtn   : BOOL;
    resetBtn   : BOOL;
    doneSensor : BOOL;
    targetVol  : REAL;
    flowVol    : REAL;
END_VAR
VAR_OUTPUT
    valveOpen  : BOOL;
    fillsToday : INT;
END_VAR
VAR
    state           : INT;       // 0=idle, 1=filling, 2=pendingConfirm
    tmp_accVol      : REAL;      // accumulated volume for current bottle
    tmp_pending     : BOOL;      // bottle waiting for doneSensor confirmation
    prev_startBtn   : BOOL;      // previous scan startBtn (power-on FALSE)
    prev_resetBtn   : BOOL;      // previous scan resetBtn (power-on FALSE)
    tmp_risingStart : BOOL;
    tmp_risingReset : BOOL;
END_VAR

// Rising edge detection
tmp_risingStart := startBtn AND NOT prev_startBtn;
tmp_risingReset := resetBtn AND NOT prev_resetBtn;

// Update previous values
prev_startBtn := startBtn;
prev_resetBtn := resetBtn;

// State machine
IF tmp_risingReset THEN
    fillsToday := 0;
    valveOpen := FALSE;
    tmp_pending := FALSE;
    tmp_accVol := 0.0;
    state := 0;
ELSE
    CASE state OF
        0: // idle
            IF tmp_risingStart THEN
                IF tmp_pending THEN
                    tmp_pending := FALSE;
                END_IF;
                tmp_accVol := flowVol;
                IF flowVol >= targetVol THEN
                    valveOpen := FALSE;
                    tmp_pending := TRUE;
                    state := 2;
                ELSE
                    valveOpen := TRUE;
                    state := 1;
                END_IF;
            END_IF;

        1: // filling
            tmp_accVol := tmp_accVol + flowVol;
            IF tmp_accVol >= targetVol THEN
                valveOpen := FALSE;
                tmp_pending := TRUE;
                state := 2;
            END_IF;

        2: // pendingConfirm
            IF tmp_risingStart THEN
                IF tmp_pending THEN
                    tmp_pending := FALSE;
                END_IF;
                tmp_accVol := flowVol;
                IF flowVol >= targetVol THEN
                    valveOpen := FALSE;
                    tmp_pending := TRUE;
                ELSE
                    valveOpen := TRUE;
                    state := 1;
                END_IF;
            ELSIF doneSensor THEN
                IF fillsToday < 32767 THEN
                    fillsToday := fillsToday + 1;
                END_IF;
                tmp_pending := FALSE;
                state := 0;
            END_IF;
    END_CASE;
END_IF;

END_FUNCTION_BLOCK

(* ---- self-medium-04.raw_candidate_01.st ---- *)
(* ENGINEERING_CONTRACT *)
(*
PUB001-PUB005: State machine (idle/filling/pending)
- valveOpen: active in filling, reset clears it, held until target reached
- fillsToday: monotonic up, reset to 0, saturates at 32767
- pendingConfirm: set when valve closes without immediate doneSensor, cleared on confirmation or reset

PUB006: startBtn rising edge triggers new bottle (only in idle or pending)
PUB007: resetBtn rising edge takes absolute priority, clears all state
PUB008: doneSensor level-triggered confirmation (checked after valve state set)
PUB009-PUB011: flowVol accumulated per scan in tmp_accVol; start scan includes its own flowVol
PUB012-PUB016: saturation behavior, no repeat count, no count while filling
*)
(* CONTRACT_RULES [] *)

FUNCTION_BLOCK FB
VAR_INPUT
    startBtn   : BOOL;
    resetBtn   : BOOL;
    doneSensor : BOOL;
    targetVol  : REAL;
    flowVol    : REAL;
END_VAR
VAR_OUTPUT
    valveOpen  : BOOL;
    fillsToday : INT;
END_VAR
VAR
    state           : INT;       // 0=idle, 1=filling, 2=pendingConfirm
    tmp_accVol      : REAL;      // accumulated volume for current bottle
    tmp_pending     : BOOL;      // bottle waiting for doneSensor confirmation
    prev_startBtn   : BOOL;      // previous scan startBtn (power-on FALSE)
    prev_resetBtn   : BOOL;      // previous scan resetBtn (power-on FALSE)
    tmp_risingStart : BOOL;
    tmp_risingReset : BOOL;
END_VAR

// Rising edge detection
tmp_risingStart := startBtn AND NOT prev_startBtn;
tmp_risingReset := resetBtn AND NOT prev_resetBtn;

// Update previous values
prev_startBtn := startBtn;
prev_resetBtn := resetBtn;

// State machine
IF tmp_risingReset THEN
    fillsToday := 0;
    valveOpen := FALSE;
    tmp_pending := FALSE;
    tmp_accVol := 0.0;
    state := 0;
ELSE
    CASE state OF
        0: // idle
            IF tmp_risingStart THEN
                IF tmp_pending THEN
                    tmp_pending := FALSE;
                END_IF;
                tmp_accVol := flowVol;
                IF flowVol >= targetVol THEN
                    valveOpen := FALSE;
                    tmp_pending := TRUE;
                    state := 2;
                ELSE
                    valveOpen := TRUE;
                    state := 1;
                END_IF;
            END_IF;

        1: // filling
            tmp_accVol := tmp_accVol + flowVol;
            IF tmp_accVol >= targetVol THEN
                valveOpen := FALSE;
                tmp_pending := TRUE;
                state := 2;
            END_IF;

        2: // pendingConfirm
            IF tmp_risingStart THEN
                IF tmp_pending THEN
                    tmp_pending := FALSE;
                END_IF;
                tmp_accVol := flowVol;
                IF flowVol >= targetVol THEN
                    valveOpen := FALSE;
                    tmp_pending := TRUE;
                ELSE
                    valveOpen := TRUE;
                    state := 1;
                END_IF;
            ELSIF doneSensor THEN
                IF fillsToday < 32767 THEN
                    fillsToday := fillsToday + 1;
                END_IF;
                tmp_pending := FALSE;
                state := 0;
            END_IF;
    END_CASE;
END_IF;

END_FUNCTION_BLOCK

(* ---- self-medium-05.candidate_01.st ---- *)
(*
ENGINEERING_CONTRACT
================================================================================
| Output/State    | Activation          | Retention        | Reset/Deactivation | Units        |
|-----------------|---------------------|------------------|---------------------|--------------|
| qualified       | Temp∈[447,453]∧Pres∈[3750,3850] | N/A (combinational) | N/A               | Boolean      |
| dataFault       | scanSeconds∉(0,10]∨Flow∉[0,90/6] | N/A (combinational) | N/A               | Boolean      |
| qualifiedTon    | enable∧qualified∧¬fault | Hold on fault/¬enable | resetBtn rising edge | tonnes (t)   |
| fuelTon         | enable∧¬fault        | Hold on fault/¬enable | resetBtn rising edge | tonnes (t)   |
| revenue         | = qualifiedTon*280  | Derived every scan  | resetBtn rising edge | yuan (元)     |
| cost            | = fuelTon*1500      | Derived every scan  | resetBtn rising edge | yuan (元)     |
| netProfit       | = revenue-cost      | Derived every scan  | N/A (may be <0)     | yuan (元)     |
--------------------------------------------------------------------------------
Priority: resetBtn rising edge > fault freeze (same-scan: reset clears accumulators)
Interval: scanSeconds ∈ (0,10] (inclusive upper bound 10.0; >10.0 is fault)
================================================================================
*)

(* CONTRACT_RULES [] *)

FUNCTION_BLOCK FB
VAR_INPUT
    enable       : BOOL;
    resetBtn     : BOOL;
    scanSeconds  : LREAL;
    steamFlow    : LREAL;
    fuelFlow     : LREAL;
    steamTemp    : LREAL;
    steamPressure: LREAL;
END_VAR
VAR_OUTPUT
    qualified    : BOOL;
    dataFault    : BOOL;
    qualifiedTon : LREAL;
    fuelTon      : LREAL;
    revenue      : LREAL;
    cost         : LREAL;
    netProfit    : LREAL;
END_VAR
VAR
    tmp_PrevResetBtn   : BOOL := FALSE;
    tmp_ResetRising    : BOOL;
    local_QualifiedTon : LREAL := 0.0;
    local_FuelTon      : LREAL := 0.0;
END_VAR

// Detect rising edge of resetBtn
tmp_ResetRising := resetBtn AND NOT tmp_PrevResetBtn;

// Data fault detection: scanSeconds not in (0,10] OR flows out of range
dataFault := (scanSeconds <= 0.0) OR (scanSeconds > 10.0)
             OR (steamFlow < 0.0) OR (steamFlow > 90.0)
             OR (fuelFlow < 0.0) OR (fuelFlow > 6.0);

// Qualified detection: closed interval [447,453] for temp and [3750,3850] for pressure
qualified := (steamTemp >= 447.0) AND (steamTemp <= 453.0)
             AND (steamPressure >= 3750.0) AND (steamPressure <= 3850.0);

// Reset: rising edge of resetBtn takes priority; clear accumulators and skip accumulation
IF tmp_ResetRising THEN
    local_QualifiedTon := 0.0;
    local_FuelTon      := 0.0;
ELSE
    // Accumulate qualified steam: only when qualified, enabled, and no fault
    IF qualified AND enable AND NOT dataFault THEN
        local_QualifiedTon := local_QualifiedTon + (steamFlow * scanSeconds / 1000.0);
    END_IF;

    // Accumulate fuel: whenever enabled and no fault (regardless of qualified status)
    IF enable AND NOT dataFault THEN
        local_FuelTon := local_FuelTon + (fuelFlow * scanSeconds / 1000.0);
    END_IF;
END_IF;

// Update outputs
qualifiedTon := local_QualifiedTon;
fuelTon      := local_FuelTon;
revenue      := qualifiedTon * 280.0;
cost         := fuelTon * 1500.0;
netProfit    := revenue - cost;

// Update previous state for next scan edge detection
tmp_PrevResetBtn := resetBtn;

END_FUNCTION_BLOCK

(* ---- self-medium-05.raw_candidate_01.st ---- *)
(*
ENGINEERING_CONTRACT
================================================================================
| Output/State    | Activation          | Retention        | Reset/Deactivation | Units        |
|-----------------|---------------------|------------------|---------------------|--------------|
| qualified       | Temp∈[447,453]∧Pres∈[3750,3850] | N/A (combinational) | N/A               | Boolean      |
| dataFault       | scanSeconds∉(0,10]∨Flow∉[0,90/6] | N/A (combinational) | N/A               | Boolean      |
| qualifiedTon    | enable∧qualified∧¬fault | Hold on fault/¬enable | resetBtn rising edge | tonnes (t)   |
| fuelTon         | enable∧¬fault        | Hold on fault/¬enable | resetBtn rising edge | tonnes (t)   |
| revenue         | = qualifiedTon*280  | Derived every scan  | resetBtn rising edge | yuan (元)     |
| cost            | = fuelTon*1500      | Derived every scan  | resetBtn rising edge | yuan (元)     |
| netProfit       | = revenue-cost      | Derived every scan  | N/A (may be <0)     | yuan (元)     |
--------------------------------------------------------------------------------
Priority: resetBtn rising edge > fault freeze (same-scan: reset clears accumulators)
Interval: scanSeconds ∈ (0,10] (inclusive upper bound 10.0; >10.0 is fault)
================================================================================
*)

(* CONTRACT_RULES [] *)

FUNCTION_BLOCK FB
VAR_INPUT
    enable       : BOOL;
    resetBtn     : BOOL;
    scanSeconds  : LREAL;
    steamFlow    : LREAL;
    fuelFlow     : LREAL;
    steamTemp    : LREAL;
    steamPressure: LREAL;
END_VAR
VAR_OUTPUT
    qualified    : BOOL;
    dataFault    : BOOL;
    qualifiedTon : LREAL;
    fuelTon      : LREAL;
    revenue      : LREAL;
    cost         : LREAL;
    netProfit    : LREAL;
END_VAR
VAR
    tmp_PrevResetBtn   : BOOL := FALSE;
    tmp_ResetRising    : BOOL;
    local_QualifiedTon : LREAL := 0.0;
    local_FuelTon      : LREAL := 0.0;
END_VAR

// Detect rising edge of resetBtn
tmp_ResetRising := resetBtn AND NOT tmp_PrevResetBtn;

// Data fault detection: scanSeconds not in (0,10] OR flows out of range
dataFault := (scanSeconds <= 0.0) OR (scanSeconds > 10.0)
             OR (steamFlow < 0.0) OR (steamFlow > 90.0)
             OR (fuelFlow < 0.0) OR (fuelFlow > 6.0);

// Qualified detection: closed interval [447,453] for temp and [3750,3850] for pressure
qualified := (steamTemp >= 447.0) AND (steamTemp <= 453.0)
             AND (steamPressure >= 3750.0) AND (steamPressure <= 3850.0);

// Reset: rising edge of resetBtn takes priority; clear accumulators and skip accumulation
IF tmp_ResetRising THEN
    local_QualifiedTon := 0.0;
    local_FuelTon      := 0.0;
ELSE
    // Accumulate qualified steam: only when qualified, enabled, and no fault
    IF qualified AND enable AND NOT dataFault THEN
        local_QualifiedTon := local_QualifiedTon + (steamFlow * scanSeconds / 1000.0);
    END_IF;

    // Accumulate fuel: whenever enabled and no fault (regardless of qualified status)
    IF enable AND NOT dataFault THEN
        local_FuelTon := local_FuelTon + (fuelFlow * scanSeconds / 1000.0);
    END_IF;
END_IF;

// Update outputs
qualifiedTon := local_QualifiedTon;
fuelTon      := local_FuelTon;
revenue      := qualifiedTon * 280.0;
cost         := fuelTon * 1500.0;
netProfit    := revenue - cost;

// Update previous state for next scan edge detection
tmp_PrevResetBtn := resetBtn;

END_FUNCTION_BLOCK

(* ---- self-medium-06.candidate_01.st ---- *)
FUNCTION_BLOCK FB
VAR_INPUT
    enable         : BOOL;
    resetBtn       : BOOL;
    sensorValid    : BOOL;
    setpoint       : REAL;
    temperature    : REAL;
    scanSeconds    : REAL;
    bias           : REAL;
END_VAR
VAR_OUTPUT
    power          : REAL;
    correction     : REAL;
    fault          : BOOL;
END_VAR
VAR
    ePrev              : REAL := 0.0;
    prevEnableAndNotFault : BOOL := FALSE;
    prevResetBtn       : BOOL := FALSE;
    historyValid       : BOOL := FALSE;
END_VAR
(* ENGINEERING_CONTRACT
+-------------------------------------------------------------------------------------+
| Output/State Group  | Activation           | Retention   | Reset/Deactivation     |
+-------------------------------------------------------------------------------------+
| power (0..100%)     | enable & !fault &    | bias+corr   | fault|!enable|reset↑   |
|                     | !rising(resetBtn)    | clamped     | (first scan only)      |
+-------------------------------------------------------------------------------------+
| correction (±30%)   | enable & !fault &    | Σ(w·c)/Σw  | fault|!enable|reset↑   |
|                     | !rising(resetBtn)    | (centroid)  | (first scan only)      |
+-------------------------------------------------------------------------------------+
| ePrev (history)     | normal differential  | held        | fault|!enable|reset↑   |
|                     | on valid non-first   | across scan | clears to 0.0          |
|                     | scans                |             |                        |
+-------------------------------------------------------------------------------------+
| de (error deriv.)   | de=0 on first scan;  | N/A         | N/A                    |
|                     | de=(e-ePrev)/scanSec |             |                        |
|                     | on valid non-first   |             |                        |
+-------------------------------------------------------------------------------------+
| fault               | !sensorValid OR      | latched     | NOT modelled (output)  |
|                     | scanSeconds<=0 OR    | until clear |                        |
|                     | scanSeconds>10       |             |                        |
+-------------------------------------------------------------------------------------+
| PUB reference: PUB001=enable, PUB002=resetBtn↑, PUB003=sensorValid, PUB004=setpoint|
|                PUB005=temperature, PUB006=scanSeconds (s), PUB007=bias             |
|                PUB008=power[0,100], PUB009=correction, PUB010=fault conditions     |
|                PUB011-015=reset behavior, PUB016-020=first-scan de=0               |
+-------------------------------------------------------------------------------------+
*)
BEGIN
    // Fault detection: PUB010
    fault := NOT sensorValid OR scanSeconds <= 0.0 OR scanSeconds > 10.0;

    // Clear outputs and history on fault, disable, or reset rising edge: PUB011, PUB012
    IF fault OR NOT enable OR (resetBtn AND NOT prevResetBtn) THEN
        power := 0.0;
        correction := 0.0;
        ePrev := 0.0;
        historyValid := FALSE;
        // Do not update prev* here; preserve for next-scan rising detection
    ELSE
        // Normal fuzzy calculation on valid scans
        VAR temp_e : REAL;
        VAR temp_de : REAL;
        VAR x, y : REAL;
        VAR xN, xZ, xP : REAL;
        VAR yN, yZ, yP : REAL;
        VAR wNN, wNZ, wNP : REAL;
        VAR wZN, wZZ, wZP : REAL;
        VAR wPN, wPZ, wPP : REAL;
        VAR wSum : REAL;
        BEGIN
            temp_e := setpoint - temperature;

            // First scan after clear: de = 0; PUB017, PUB020
            IF NOT (prevEnableAndNotFault AND NOT (resetBtn AND NOT prevResetBtn)) THEN
                // First scan or history was cleared
                temp_de := 0.0;
                historyValid := FALSE;
            ELSE
                // Normal differential: PUB019
                IF scanSeconds > 0.0 THEN
                    temp_de := (temp_e - ePrev) / scanSeconds;
                ELSE
                    temp_de := 0.0;
                END_IF;
                historyValid := TRUE;
            END_IF;

            // Normalize: x = clamp(e/10, -1, 1), y = clamp(de/2, -1, 1); PUB005
            x := temp_e / 10.0;
            IF x > 1.0 THEN x := 1.0; ELSIF x < -1.0 THEN x := -1.0; END_IF;
            y := temp_de / 2.0;
            IF y > 1.0 THEN y := 1.0; ELSIF y < -1.0 THEN y := -1.0; END_IF;

            // Membership functions: μN(z)=max(-z,0), μZ(z)=1-|z|, μP(z)=max(z,0); PUB003
            xN := 0.0; IF x < 0.0 THEN xN := -x; END_IF;
            xZ := 1.0 - ABS(x); IF xZ < 0.0 THEN xZ := 0.0; END_IF;
            xP := 0.0; IF x > 0.0 THEN xP := x; END_IF;

            yN := 0.0; IF y < 0.0 THEN yN := -y; END_IF;
            yZ := 1.0 - ABS(y); IF yZ < 0.0 THEN yZ := 0.0; END_IF;
            yP := 0.0; IF y > 0.0 THEN yP := y; END_IF;

            // Rule weights: w(i,j) = μi(x) × μj(y); PUB004
            wNN := xN * yN;
            wNZ := xN * yZ;
            wNP := xN * yP;
            wZN := xZ * yN;
            wZZ := xZ * yZ;
            wZP := xZ * yP;
            wPN := xP * yN;
            wPZ := xP * yZ;
            wPP := xP * yP;

            // Centroid defuzzification: correction = Σ(w·c)/Σw; PUB004
            wSum := wNN + wNZ + wNP + wZN + wZZ + wZP + wPN + wPZ + wPP;
            IF wSum > 0.0 THEN
                correction := (wNN * (-30.0) + wNZ * (-20.0) + wNP * (-10.0) +
                               wZN * (-10.0) + wZZ *   0.0 + wZP *   10.0 +
                               wPN *  10.0 + wPZ *   20.0 + wPP *   30.0) / wSum;
            ELSE
                correction := 0.0;
            END_IF;

            // Update ePrev for next scan: PUB018
            ePrev := temp_e;
        END;

        // Power: clamp(bias + correction, 0, 100); correction NOT clamped; PUB009
        power := bias + correction;
        IF power > 100.0 THEN power := 100.0;
        ELSIF power < 0.0 THEN power := 0.0;
        END_IF;
    END_IF;

    // Update state tracking for next scan; PUB002 (rising edge detection)
    prevEnableAndNotFault := enable AND NOT fault;
    prevResetBtn := resetBtn;
END_FUNCTION_BLOCK
